(* IEC 61131-3 sources: trust-platform/examples/control/01-feedback-foundations-and-temperature-control/11-measurement-filtering/src, 2 files *)

(* ---- Main.st ---- *)
USING Control;

(* Fraction of the raw-minus-filtered difference applied per update: alpha = dt/(Tf + dt). *)
FUNCTION FilterFraction : LREAL
VAR_INPUT
    CycleTime : LREAL;
    FilterTime : LREAL;
END_VAR
FilterFraction := CycleTime / (FilterTime + CycleTime);
END_FUNCTION

(* First-order low-pass update: yf_new = yf_old + alpha·(yr − yf_old). *)
FUNCTION FilterUpdate : LREAL
VAR_INPUT
    PreviousFilteredValue : LREAL;
    RawValue : LREAL;
    FilterFraction : LREAL;
END_VAR
FilterUpdate := PreviousFilteredValue + FilterFraction * (RawValue - PreviousFilteredValue);
END_FUNCTION

(* Proportional request around the holding output: u = u_hold + Kp·(SP − measurement). *)
FUNCTION ProportionalRequest : LREAL
VAR_INPUT
    HoldingOutput : LREAL;
    ProportionalGain : LREAL;
    Setpoint : LREAL;
    Measurement : LREAL;
END_VAR
ProportionalRequest := HoldingOutput + ProportionalGain * (Setpoint - Measurement);
END_FUNCTION

FUNCTION SamePidParameters : BOOL
VAR_INPUT
    Left : Control.PIDParameters;
    Right : Control.PIDParameters;
END_VAR
SamePidParameters :=
    Left.ProportionalGain = Right.ProportionalGain
    AND Left.IntegralGain = Right.IntegralGain
    AND Left.DerivativeGain = Right.DerivativeGain
    AND Left.ProportionalSetpointWeight = Right.ProportionalSetpointWeight
    AND Left.DerivativeSetpointWeight = Right.DerivativeSetpointWeight
    AND Left.Bias = Right.Bias
    AND Left.OutputMinimum = Right.OutputMinimum
    AND Left.OutputMaximum = Right.OutputMaximum
    AND Left.RateMinimum = Right.RateMinimum
    AND Left.RateMaximum = Right.RateMaximum
    AND Left.TrackingTime = Right.TrackingTime
    AND Left.AntiWindup = Right.AntiWindup;
END_FUNCTION

PROGRAM Main
VAR
    Controller : Control.PID;
    (* Tune replaces this record with each candidate; the defaults are the Lesson 23
       controller: the relay gains with the setpoint weight 0.3 applied there. *)
    Parameters : Control.PIDParameters := (
        ProportionalGain := LREAL#13.0,
        IntegralGain := LREAL#3.5,
        DerivativeGain := LREAL#0.0,
        ProportionalSetpointWeight := LREAL#0.3,
        DerivativeSetpointWeight := LREAL#0.0,
        Bias := LREAL#0.0,
        OutputMinimum := LREAL#0.0,
        OutputMaximum := LREAL#100.0,
        RateMinimum := LREAL#-10000.0,
        RateMaximum := LREAL#10000.0,
        TrackingTime := LREAL#1.0,
        AntiWindup := PIDAntiWindup#BackCalculation
    );
    ConfiguredParameters : Control.PIDParameters;
    ParameterRevision : DINT := 0;
    InitialState : Control.PIDInitialState;
    ObservedState : Control.PIDInitialState;
    Input : Control.PIDInput;
    Initialized : BOOL := FALSE;
    AutoMode : BOOL := FALSE;
    ManualOutput : LREAL := 75.0;
    SafetyAbort : BOOL := FALSE;
    DataUsable : BOOL := FALSE;
    SetpointC : LREAL := 35.0;
    DisturbanceKw : LREAL := 0.0;
    WaterInputC : LREAL := 35.0;
    WaterTemperatureC : LREAL := 35.0;
    TemperatureC : LREAL := 35.0;
    SafeProcessValueC : LREAL := 35.0;
    AppliedPowerPct : LREAL := 75.0;
    RequestedPowerPct : LREAL := 75.0;
    ErrorC : LREAL := 0.0;
    (* Reference of the weighted proportional term: the 35 °C hot operating point. *)
    OperatingPointC : LREAL := 35.0;
    (* Measurement filter: Tf = 0 bypasses it; Control Studio applies Tf with the gains. *)
    FilterTimeS : LREAL := 0.0;
    FilterAlpha : LREAL := 1.0;
    FilteredC : LREAL := 35.0;
    FilterActive : BOOL := FALSE;
    FilterWasActive : BOOL := FALSE;
    ProportionalPct : LREAL := 0.0;
    IntegralPct : LREAL := 75.0;
    PreviousAppliedPct : LREAL := 75.0;
    CommandActivityPoints : LREAL := 0.0;
END_VAR

(* The Lesson 21 heater: both feedback bindings observe the heated water, and the
   temperature measurement carries ±0.02 °C noise. The controller uses the filtered value. *)
WaterTemperatureC := WaterInputC;
DataUsable := TemperatureC >= LREAL#0.0 AND TemperatureC <= LREAL#80.0;
IF DataUsable THEN
    SafeProcessValueC := TemperatureC;
ELSE
    SafetyAbort := TRUE;
END_IF;
(* Tf = 0 gives alpha = 1: the filtered value equals the raw measurement (bypass). *)
FilterAlpha := FilterFraction(CycleTime := LREAL#0.1, FilterTime := MAX(FilterTimeS, LREAL#0.0));

(* Control Studio's Apply replaces this complete record at the task boundary; the
   program copies it into the actual controller and never overwrites it cyclically. *)
IF NOT Initialized OR NOT SamePidParameters(Left := Parameters, Right := ConfiguredParameters) THEN
    ConfiguredParameters := Parameters;
    ParameterRevision := ParameterRevision + 1;
END_IF;
Controller.Configure(Parameters := Parameters);

IF NOT Initialized THEN
    (* Common hot reset: the heater already holds 35 °C with 75 % output, so the
       controller's retained output starts at the holding command. *)
    ManualOutput := LREAL#75.0;
    IF NOT AutoMode THEN
        SetpointC := SafeProcessValueC;
    END_IF;
    FilteredC := SafeProcessValueC;
    InitialState.Setpoint := SetpointC;
    InitialState.ProcessValue := SafeProcessValueC;
    InitialState.NominalOutput := ManualOutput;
    InitialState.SaturatedOutput := ManualOutput;
    InitialState.SetpointRate := LREAL#0.0;
    InitialState.ProcessValueRate := LREAL#0.0;
    InitialState.FeedForward := LREAL#0.0;
    Controller.Initialize(State := InitialState);
    Initialized := TRUE;
END_IF;

(* The filter runs while the controller is in Auto. In Manual and in the Auto-entry scan it
   restarts from the fresh measurement, the value the transfer aligned the controller to, so
   entering Auto is exactly bumpless; filtering starts with the next scan. *)
FilterActive := AutoMode AND NOT SafetyAbort AND Parameters.ProportionalGain > LREAL#0.0
    AND Parameters.IntegralGain > LREAL#0.0;
IF Initialized AND FilterActive AND FilterWasActive THEN
    FilteredC := FilterUpdate(PreviousFilteredValue := FilteredC, RawValue := SafeProcessValueC, FilterFraction := FilterAlpha);
ELSE
    FilteredC := SafeProcessValueC;
END_IF;
FilterWasActive := FilterActive;
Input.Setpoint := SetpointC;
Input.ProcessValue := FilteredC;
Input.CycleTime := LREAL#0.1;
Input.FeedForward := LREAL#0.0;
Input.TrackingOutput := ManualOutput;
IF SafetyAbort THEN
    (* An abort or invalid measurement removes heat and the test load until a full restart. *)
    Input.Mode := PIDMode#Manual;
    Input.ManualOutput := LREAL#0.0;
    DisturbanceKw := LREAL#0.0;
ELSIF AutoMode AND Parameters.ProportionalGain > LREAL#0.0 AND Parameters.IntegralGain > LREAL#0.0 THEN
    Input.Mode := PIDMode#Auto;
    Input.ManualOutput := ManualOutput;
ELSE
    Input.Mode := PIDMode#Manual;
    Input.ManualOutput := ManualOutput;
END_IF;
ErrorC := SetpointC - FilteredC;
AppliedPowerPct := Controller.Update(Input := Input);

(* Diagnostics come from the actual controller state; the PI equations live in Control.PID.
   Command activity adds every applied-command movement, starting from the 75% holding command. *)
ObservedState := Controller.GetState();
RequestedPowerPct := ObservedState.NominalOutput;
IF Input.Mode = PIDMode#Auto THEN
    (* Weighted P = Kp·(β·(SP − T0) − (PV − T0)); the integral uses the full error. *)
    ProportionalPct := Parameters.ProportionalGain * (Parameters.ProportionalSetpointWeight * (SetpointC - OperatingPointC)
        - (FilteredC - OperatingPointC));
ELSE
    ProportionalPct := LREAL#0.0;
END_IF;
IntegralPct := RequestedPowerPct - ProportionalPct;
CommandActivityPoints := CommandActivityPoints + ABS(AppliedPowerPct - PreviousAppliedPct);
PreviousAppliedPct := AppliedPowerPct;

END_PROGRAM

CONFIGURATION Config
RESOURCE Res ON PLC
    TASK MainTask(INTERVAL := T#100ms, PRIORITY := 1);
    PROGRAM P1 WITH MainTask : Main;
END_RESOURCE
VAR_CONFIG
    P1.SafetyAbort AT %MX96.3 : BOOL;
    P1.DataUsable AT %MX96.2 : BOOL;
    P1.AppliedPowerPct AT %QL0 : LREAL;
    P1.DisturbanceKw AT %QL8 : LREAL;
    P1.WaterInputC AT %IL0 : LREAL;
    P1.TemperatureC AT %IL8 : LREAL;
    P1.SetpointC AT %ML0 : LREAL;
    P1.IntegralPct AT %ML16 : LREAL;
    P1.RequestedPowerPct AT %ML32 : LREAL;
    P1.WaterTemperatureC AT %ML48 : LREAL;
    P1.ProportionalPct AT %ML56 : LREAL;
    P1.CommandActivityPoints AT %ML64 : LREAL;
    P1.ManualOutput AT %ML72 : LREAL;
END_VAR
END_CONFIGURATION

(* ---- tests.st ---- *)
(* @trustlsp:runtime-ignore — run these assertions with trust-dev test;
   they are not scheduled PLC instances in the lesson simulator. *)
TEST_PROGRAM FilterMovesPartwayTowardRawMeasurement
VAR
    Fraction : LREAL;
    Filtered : LREAL;
END_VAR
Fraction := FilterFraction(CycleTime := LREAL#0.1, FilterTime := LREAL#1.0);
Filtered := FilterUpdate(PreviousFilteredValue := LREAL#35.0, RawValue := LREAL#36.0, FilterFraction := Fraction);
ASSERT_NEAR(EXPECTED := LREAL#0.0909090909090909, ACTUAL := Fraction, DELTA := LREAL#1.0e-12);
ASSERT_NEAR(EXPECTED := LREAL#35.0909090909091, ACTUAL := Filtered, DELTA := LREAL#1.0e-12);
END_TEST_PROGRAM

TEST_PROGRAM FilteredMeasurementReducesRequestMovement
VAR
    RawRequest : LREAL;
    FilteredRequest : LREAL;
END_VAR
RawRequest := ProportionalRequest(HoldingOutput := LREAL#75.0, ProportionalGain := LREAL#2.0, Setpoint := LREAL#35.0, Measurement := LREAL#36.0);
FilteredRequest := ProportionalRequest(HoldingOutput := LREAL#75.0, ProportionalGain := LREAL#2.0, Setpoint := LREAL#35.0, Measurement := LREAL#35.0909090909091);
ASSERT_TRUE(IN := RawRequest = LREAL#73.0);
ASSERT_NEAR(EXPECTED := LREAL#74.8181818181818, ACTUAL := FilteredRequest, DELTA := LREAL#1.0e-12);
END_TEST_PROGRAM
